DATA_BLOCK "GDB_LineOwnerTest"
{ S7_Optimized_Access := 'TRUE' }
VERSION : 0.1
NON_RETAIN
VAR
    PoisonPulse : Bool;
    Poisoned {ExternalWritable := 'False'} : Bool;
    BootDefaultSeen {ExternalWritable := 'False'} : Bool;
    BootDefaultValue {ExternalWritable := 'False'} : UDInt;
    WorkingTaktMs {ExternalWritable := 'False'} : UDInt;
END_VAR
BEGIN
END_DATA_BLOCK
